(* IEC 61131-3 sources: plc-process-lib/tests/DUTs/TestDevice, 4 files *)

(* ---- ST_TestDeviceCfg.dut.st ---- *)
// Назначение: конфигурация тестового устройства FB_TestDevice. Заканчивается полями тревог, как
//             ST_<Dev>Cfg библиотеки (udiAlarmIdBase, astAlarm). Значения по умолчанию проходят
//             CheckConfig. Только для тестов.
// Автор:      kr0nsch
// Версия:     0.1.0
// Документ:   docs/TESTING.md, раздел «Тестовое устройство»
{attribute 'qualified_only'}
TYPE ST_TestDeviceCfg :
STRUCT
    rGain          : REAL := 2.0;    // коэффициент; корректен, если конечен и > 0 (бит 0 wCfgErr)
    tRunDelay      : TIME := T#0S;   // задержка включения в Auto (вложенный FB_Delay до BeginCycle)
    udiAlarmIdBase : UDINT := 0;     // номер первой тревоги устройства
    astAlarm       : ARRAY[0..GVL_Const.DEV_ALARMS_MAX - 1] OF ST_AlarmCfg;   // по слотам; умолчания ST_AlarmCfg
END_STRUCT
END_TYPE

(* ---- ST_TestDeviceCmd.dut.st ---- *)
// Назначение: команды тестового устройства FB_TestDevice — общий заголовок и команды механизма,
//             как у ST_<Dev>Cmd библиотеки. Только для тестов.
// Автор:      kr0nsch
// Версия:     0.1.0
// Документ:   docs/TESTING.md, раздел «Тестовое устройство»
{attribute 'qualified_only'}
TYPE ST_TestDeviceCmd :
STRUCT
    stCommon : ST_DeviceCmd;   // общий заголовок
    xStart   : BOOL;           // импульс: пуск (Manual)
    xStop    : BOOL;           // импульс: стоп (в Auto — переход в Manual и стоп)
    uiTrace  : UINT;           // пишет тело наследника FB_TestDeviceExt после SUPER^ (проверка R3)
END_STRUCT
END_TYPE

(* ---- ST_TestDeviceSts.dut.st ---- *)
// Назначение: состояние тестового устройства FB_TestDevice: общий заголовок и значение по LKG.
//             Только для тестов.
// Автор:      kr0nsch
// Версия:     0.1.0
// Документ:   docs/TESTING.md, раздел «Тестовое устройство»
{attribute 'qualified_only'}
TYPE ST_TestDeviceSts :
STRUCT
    stCommon : ST_DeviceSts;   // общий заголовок
    rOut_eu  : REAL;           // значение по конфигурации LKG: rGain * 10
END_STRUCT
END_TYPE

(* ---- U_TestEnumInt.dut.st ---- *)
// Назначение: значение вне строгого перечисления для тестов санитизации. Строгое перечисление не
//             даёт присвоить число в исходном тексте (C0358), а в памяти persistent оно может быть
//             любым: тест пишет iValue и читает поле перечисления. Только для тестов.
// Автор:      kr0nsch
// Версия:     0.1.0
// Документ:   docs/TESTING.md, раздел «Тестовое устройство»
{attribute 'qualified_only'}
TYPE U_TestEnumInt :
UNION
    iValue    : INT;               // число, которое пишет тест
    eMode     : E_DeviceMode;      // то же как режим
    ePriority : E_AlarmPriority;   // то же как приоритет тревоги
END_UNION
END_TYPE
